TYPE T_MotorName : STRING(40);
END_TYPE

(* stored: Version 1.1.0.1
   DUT T_MotorName: Id {f31eddd5-f155-472f-bbd3-fa1b1a381526} *)
